(* IEC 61131-3 sources: volt/packages/volt-lsp-iec/test-corpus/lenze-mid/Device/Plc Logic/Application/Library Manager/CmpDynamicText, 22 files *)

(* ---- DYNAMICTEXTCHANGELANGUAGE.pou ---- *)
FUNCTION DYNAMICTEXTCHANGELANGUAGE : BOOL
VAR_INPUT
	STLANGUAGE : STRING;
END_VAR
END_FUNCTION

(* ---- DYNAMICTEXTGETCURRENTLANGUAGE.pou ---- *)
FUNCTION DYNAMICTEXTGETCURRENTLANGUAGE : STRING
END_FUNCTION

(* ---- DYNAMICTEXTGETDEFAULTTEXT.pou ---- *)
FUNCTION DYNAMICTEXTGETDEFAULTTEXT : POINTER TO STRING
VAR_INPUT
	PSTTEXTLIST : POINTER TO STRING;
	PSTTEXTINDEX : POINTER TO STRING;
END_VAR
END_FUNCTION

(* ---- DYNAMICTEXTGETDEFAULTTEXTW.pou ---- *)
FUNCTION DYNAMICTEXTGETDEFAULTTEXTW : POINTER TO STRING
VAR_INPUT
	PSTTEXTLIST : POINTER TO STRING;
	PSTTEXTINDEX : POINTER TO STRING;
END_VAR
END_FUNCTION

(* ---- DYNAMICTEXTGETLANGUAGETEXT.pou ---- *)
FUNCTION DYNAMICTEXTGETLANGUAGETEXT : POINTER TO STRING
VAR_IN_OUT
	STLANGUAGE : STRING;
	STTEXTLIST : STRING;
	STTEXTINDEX : STRING;
END_VAR
END_FUNCTION

(* ---- DYNAMICTEXTGETLANGUAGETEXTW.pou ---- *)
FUNCTION DYNAMICTEXTGETLANGUAGETEXTW : POINTER TO WSTRING
VAR_IN_OUT
	STLANGUAGE : STRING;
	STTEXTLIST : STRING;
	STTEXTINDEX : STRING;
END_VAR
END_FUNCTION

(* ---- DYNAMICTEXTGETTEXT.pou ---- *)
FUNCTION DYNAMICTEXTGETTEXT : POINTER TO STRING
VAR_INPUT
	PSTTEXTLIST : POINTER TO STRING;
	PSTTEXTINDEX : POINTER TO STRING;
END_VAR
END_FUNCTION

(* ---- DYNAMICTEXTGETTEXTW.pou ---- *)
FUNCTION DYNAMICTEXTGETTEXTW : POINTER TO STRING
VAR_INPUT
	PSTTEXTLIST : POINTER TO STRING;
	PSTTEXTINDEX : POINTER TO STRING;
END_VAR
END_FUNCTION

(* ---- DYNAMICTEXTITERATEINDICES.pou ---- *)
FUNCTION DYNAMICTEXTITERATEINDICES : RTS_IEC_RESULT
VAR_INPUT
	PSTTEXTLIST : POINTER TO STRING;
	PFITERATIONCALLBACK : POINTER TO BYTE;
	ITERATIONDATA : __UXINT;
END_VAR
END_FUNCTION

(* ---- DYNAMICTEXTITERATELANGUAGES.pou ---- *)
FUNCTION DYNAMICTEXTITERATELANGUAGES : RTS_IEC_RESULT
VAR_INPUT
	PFITERATIONCALLBACK : POINTER TO BYTE;
	ITERATIONDATA : __UXINT;
END_VAR
END_FUNCTION

(* ---- DYNAMICTEXTLOADDEFAULTTEXTS.pou ---- *)
FUNCTION DYNAMICTEXTLOADDEFAULTTEXTS : RTS_IEC_RESULT
END_FUNCTION

(* ---- DYNAMICTEXTLOADLANGUAGE.pou ---- *)
FUNCTION DYNAMICTEXTLOADLANGUAGE : RTS_IEC_RESULT
VAR_INPUT
	STLANGUAGE : STRING;
END_VAR
END_FUNCTION

(* ---- DYNAMICTEXTREGISTERFILE.pou ---- *)
FUNCTION DYNAMICTEXTREGISTERFILE : RTS_IEC_RESULT
VAR_INPUT
	SZFILE : REFERENCE TO STRING;
END_VAR
END_FUNCTION

(* ---- DYNAMICTEXTREGISTERPATH.pou ---- *)
FUNCTION DYNAMICTEXTREGISTERPATH : RTS_IEC_RESULT
VAR_INPUT
	SZPATH : REFERENCE TO STRING;
END_VAR
END_FUNCTION

(* ---- DYNAMICTEXTRELEASELANGUAGES.pou ---- *)
FUNCTION DYNAMICTEXTRELEASELANGUAGES : RTS_IEC_RESULT
VAR_INPUT
	XFORCERELEASE : BOOL;
END_VAR
END_FUNCTION

(* ---- DYNAMICTEXTRELEASELOCK.pou ---- *)
FUNCTION DYNAMICTEXTRELEASELOCK : BOOL
END_FUNCTION

(* ---- DYNAMICTEXTRELOADTEXTS.pou ---- *)
FUNCTION DYNAMICTEXTRELOADTEXTS : RTS_IEC_RESULT
END_FUNCTION

(* ---- DYNAMICTEXTSETLOCK.pou ---- *)
FUNCTION DYNAMICTEXTSETLOCK : BOOL
END_FUNCTION

(* ---- DYNAMICTEXTTESTANDSETLOCK.pou ---- *)
FUNCTION DYNAMICTEXTTESTANDSETLOCK : BOOL
END_FUNCTION

(* ---- DYNAMICTEXTUNLOADLANGUAGE.pou ---- *)
FUNCTION DYNAMICTEXTUNLOADLANGUAGE : RTS_IEC_RESULT
VAR_INPUT
	STLANGUAGE : STRING;
END_VAR
END_FUNCTION

(* ---- DYNAMICTEXTUNREFERENCELANGUAGE.pou ---- *)
FUNCTION DYNAMICTEXTUNREFERENCELANGUAGE : RTS_IEC_RESULT
VAR_INPUT
	STLANGUAGE : STRING;
END_VAR
END_FUNCTION

(* ---- DYNAMICTEXTUNREGISTERFILE.pou ---- *)
FUNCTION DYNAMICTEXTUNREGISTERFILE : RTS_IEC_RESULT
VAR_INPUT
	SZFILE : REFERENCE TO STRING;
END_VAR
END_FUNCTION
